(* IEC 61131-3 sources: rusty/tests/lit/single/control_statements/for_unsigned_counter, 7 files *)

(* ---- dword_counter_across_midpoint.st ---- *)
// RUN: %COMPILE %s && %RUN | %CHECK %s
//
// A FOR loop with a DWORD counter runs through the midpoint 2^31 like through any other value.

FUNCTION main
    VAR
        i : DWORD;
        first : DWORD := 16#7FFF_FFFE;
        last : DWORD := 16#8000_0001;
    END_VAR
    FOR i := first TO last DO
        printf('%u$N', i);
    END_FOR
    // CHECK:      2147483646
    // CHECK-NEXT: 2147483647
    // CHECK-NEXT: 2147483648
    // CHECK-NEXT: 2147483649
    // CHECK-NOT:  {{.+}}
END_FUNCTION

(* ---- udint_bounds_from_variables.st ---- *)
// RUN: %COMPILE %s && %RUN | %CHECK %s
//
// A FOR loop with a UDINT counter and UDINT bound variables compares the counter with the end as
// unsigned values, so it runs through the midpoint 2^31.

FUNCTION main
    VAR
        i : UDINT;
        first : UDINT := 16#7FFF_FFFE;
        last : UDINT := 16#8000_0001;
    END_VAR
    FOR i := first TO last DO
        printf('%u$N', i);
    END_FOR
    // CHECK:      2147483646
    // CHECK-NEXT: 2147483647
    // CHECK-NEXT: 2147483648
    // CHECK-NEXT: 2147483649
    // CHECK-NOT:  {{.+}}
END_FUNCTION

(* ---- udint_counter_across_midpoint.st ---- *)
// RUN: %COMPILE %s && %RUN | %CHECK %s
//
// A FOR loop with a UDINT counter runs through the midpoint 2^31 like through any other value.

FUNCTION main
    VAR
        i : UDINT;
    END_VAR
    FOR i := 16#7FFF_FFFE TO 16#8000_0001 DO
        printf('%u$N', i);
    END_FOR
    // CHECK:      2147483646
    // CHECK-NEXT: 2147483647
    // CHECK-NEXT: 2147483648
    // CHECK-NEXT: 2147483649
    // CHECK-NOT:  {{.+}}
END_FUNCTION

(* ---- udint_counter_counting_down.st ---- *)
// RUN: %COMPILE %s && %RUN | %CHECK %s
//
// A FOR loop with a UDINT counter and a negative step counts down through the midpoint 2^31.

FUNCTION main
    VAR
        i : UDINT;
    END_VAR
    FOR i := 16#8000_0001 TO 16#7FFF_FFFE BY -1 DO
        printf('%u$N', i);
    END_FOR
    // CHECK:      2147483649
    // CHECK-NEXT: 2147483648
    // CHECK-NEXT: 2147483647
    // CHECK-NEXT: 2147483646
    // CHECK-NOT:  {{.+}}
END_FUNCTION

(* ---- udint_end_from_subtraction.st ---- *)
// RUN: %COMPILE %s && %RUN | %CHECK %s
//
// `FOR i := 0 TO count - 1` with a UDINT counter and `count = 0` runs zero times, because
// `count - 1` runs in DINT and is -1.

FUNCTION main
    VAR
        i : UDINT;
        count : UDINT := 0;
        passes : DINT := 0;
    END_VAR
    FOR i := 0 TO count - 1 DO
        passes := passes + 1;
        IF passes >= 3 THEN
            EXIT;
        END_IF
    END_FOR
    printf('passes: %d$N', passes);
    // CHECK: passes: 0
END_FUNCTION

(* ---- udint_step_from_variable.st ---- *)
// RUN: %COMPILE %s && %RUN | %CHECK %s
//
// A FOR loop with a UDINT counter and a UDINT step variable runs through the midpoint 2^31.

FUNCTION main
    VAR
        i : UDINT;
        first : UDINT := 16#7FFF_FFFE;
        last : UDINT := 16#8000_0002;
        step : UDINT := 2;
    END_VAR
    FOR i := first TO last BY step DO
        printf('%u$N', i);
    END_FOR
    // CHECK:      2147483646
    // CHECK-NEXT: 2147483648
    // CHECK-NEXT: 2147483650
    // CHECK-NOT:  {{.+}}
END_FUNCTION

(* ---- ulint_counter_across_midpoint.st ---- *)
// RUN: %COMPILE %s && %RUN | %CHECK %s
//
// A FOR loop with a ULINT counter runs through the midpoint 2^63 like through any other value.

FUNCTION main
    VAR
        i : ULINT;
        first : ULINT := 16#7FFF_FFFF_FFFF_FFFE;
        last : ULINT := 16#8000_0000_0000_0001;
    END_VAR
    FOR i := first TO last DO
        printf('%llu$N', i);
    END_FOR
    // CHECK:      9223372036854775806
    // CHECK-NEXT: 9223372036854775807
    // CHECK-NEXT: 9223372036854775808
    // CHECK-NEXT: 9223372036854775809
    // CHECK-NOT:  {{.+}}
END_FUNCTION
